FUNCTION_BLOCK Heat_Control (* Composite Function Block Type *)
  (* Standard: 61499-2 *)
  (* Version 0.0, 1/6/2020, prana, nxtControl GmbH, template *)
  PACKAGE Main;
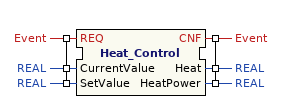
  EVENT_INPUT
    REQ WITH CurrentValue, SetValue; (* Normal Execution Request *)
  END_EVENT
  EVENT_OUTPUT
    CNF WITH Heat, HeatPower; (* Execution Confirmation *)
  END_EVENT
  VAR_INPUT
    CurrentValue : REAL; (* Input event qualifier *)
    SetValue : REAL;
  END_VAR
  VAR_OUTPUT
    Heat : REAL;
    HeatPower : REAL;
  END_VAR
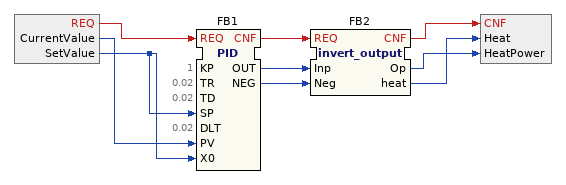
  FBS
    FB1 : PID(KP := 1, TR := 0.02, TD := 0.02, DLT := 0.02);
    FB2 : invert_output;
  END_FBS
  EVENT_CONNECTIONS
    FB2.CNF TO CNF;
    REQ TO FB1.REQ;
    FB1.CNF TO FB2.REQ;
  END_CONNECTIONS
  DATA_CONNECTIONS
    FB2.heat TO Heat;
    CurrentValue TO FB1.PV;
    SetValue TO FB1.SP;
    SetValue TO FB1.X0;
    FB1.OUT TO FB2.Inp;
    FB1.NEG TO FB2.Neg;
    FB2.Op TO HeatPower;
  END_CONNECTIONS
END_FUNCTION_BLOCK
